(* IEC 61131-3 sources: Lasal-MCP/examples/SampleSource/LASALScreenAdvancedSolution/LASALScreenAdvancedSolution/LASALScreenAdvacnedSolution/Stations/MachineControl/MachineControl/Class/VaranManager (part 4) *)

      //look in all peripheral sync outs
      for i := 1 to VM_MAX_SYNC_OUTS - 1 do

        //look if sync out id is correct
        if ( p_SyncOut^.ucSyncOutID = VM_SYNC_OUT_ID ) then

          //if it is right pll for right manager number (first is vor VaranManager number 0, second for VaranManager number 1, ....)
          if ( ud_counter = 0 ) then
            exit;					//we found right sync out --> exit
          end_if;
          ud_counter -= 1;			//we find one for lower VaranManager number
        end_if;

        //get pointer to next sync out
        p_SyncOut += sizeof ( LSL_VARANPLLSYNCOUT );

        //if we searched all sync outs set VaranManager off
        if ( i = VM_MAX_SYNC_OUTS - 1 ) then
          p_SyncOut := NIL;
          State 		:= _NotInitialized;
          ManagerOn	:= 0;
          return;
        end_if;
      end_for;

      //disable varan manager sync out
      p_SyncOut^.ucControlStatus := 0;
    end_if;

  else // if b_PayloadSupport ****************************************************************************

    // if there is no VARAN Interface available, we would crash at the call
    if pVaran = NIL then
      sd_retval := VARANMANAGER_DRIVER_NOT_EXISTS;
      return;
    end_if;

      //-----------------------------------------------------------------------------------------------
    //get manager node info from os
    ManagerNodeString := 0;

    //call OS - function (must be OS-funciton because of error handling)
    sd_retval := VARAN_iGetNodeInfo	( uiManager	:= VaranManagerNr
                                    , pucNode	  := #ManagerNodeString
                                    , pNodeInfo	:= #p_NodeInfo
                                    );

    if	( sd_retval <> VARANMANAGER_OK
      | p_NodeInfo = NIL
      )
    then
      State := _NoHardware;
      return;
    end_if;

      // get release of FPGA
    Release := p_NodeInfo^.ucFPGAVersion;

    //-----------------------------------------------------------------------------------------------
    //get Manager structure
    sd_retval := VARAN_iGetManagerControl	( uiManager := VaranManagerNr
                                          , pvCB 		  := ( #p_ManagerStructure )$^PLSL_CONTROLBLOCK
                                          , pvPLL		  := ( #p_ManagerPll )$^PLSL_VARANPLL
                                          );

    //look for an error
    if	( sd_retval 			<> 	VARANMANAGER_OK
      | p_ManagerStructure	=	NIL
      | p_ManagerPll			= 	NIL
      )
    then
      State 		:= _NotInitialized;
      ManagerOn	:= 0;
      return;
    end_if;

    //look for right sync out pointer
    p_SyncOut := #p_ManagerPll^.sSynOutPeripheral1;
    ud_Counter := VaranManagerNr;

    //look in all peripheral sync outs
    for i := 1 to VM_MAX_SYNC_OUTS - 1 do

      //look if sync out id is correct
      if ( p_SyncOut^.ucSyncOutID = VM_SYNC_OUT_ID ) then

        //if it is right pll for right manager number (first is for VaranManager number 0, second for VaranManager number 1, ....)
        if ( ud_counter = 0 ) then
          exit;					//we found right sync out --> exit
        end_if;
        ud_counter -= 1;			//we find one for lower VaranManager number
      end_if;

      //get pointer to next sync out
      p_SyncOut += sizeof ( LSL_VARANPLLSYNCOUT );

      //if we searched all sync outs set VaranManager off
      if ( i = VM_MAX_SYNC_OUTS - 1 ) then
        p_SyncOut := NIL;
        State 		:= _NotInitialized;
        ManagerOn	:= 0;
        return;
      end_if;
    end_for;

    //disable varan manager sync out
    p_SyncOut^.ucControlStatus := 0;

    //set required bit on (for varan error in init (os set bit in function InitApp) later)
    p_ManagerStructure^.ucTCEnable := p_ManagerStructure^.ucTCEnable or 16#80;

    //Get ISO start Time
    GetISOStartTime();

    p_ManagerStructure^.uiIsoStartPoint := VaranManagerTime * IsoStartPoint / 100;

  end_if; // if b_PayloadSupport ****************************************************************************

  // get maintimer in ns to compare with varan times
  MainTimer := _ClockTicks * 1000;

  //look if VaranManagerTime is a multiple of maintimer (maintimer has to be always less or equal the varan time)
  if ( VaranManagerTime mod MainTimer <> 0 ) then
    //Log entry
#ifdef HWC_LogValue2
    HWC_LogValue2(this, "@064A (VaranManager::FirstInit) VaranManagerTime ({0}) is not a multiple of MainTimer ({1})!", VaranManagerTime, MainTimer);
#endif

    State 		:= _NotInitialized;
    ManagerOn	:= 0;
    return;
  end_if;

//------------------------------------------------------------ Client Instructions --------------------------------------------------------|
//                                                                                                                                         V
  if ( IsAlsoClient ) then

    if b_PayloadSupport &
       pMultiVaran^.udVersion >= VM_MULTIVARAN_VERSION_FULL_PAYLOAD_AVAILABLE  then
      sd_retval := MULTI_VARAN_iGetNodeProperty(  hNodeHandle       := vmNodeHandle
                                                , udPropertyId      := VC_OPT_PROP_BUFFER_ADDRESS_ISO // = Offset 0 in p_ManagerClientSpace
                                                , pudPropertyValue  := (#p_ManagerClientSpace)$^UDINT );

    elsif ( _RTOSVersion >= 16#11DA ) & pVaran then

      //Schnittstelle vom OS holen!!!!!!
      sd_retval := VARAN_iGetManagerClientAddress	( uiManager		:= VaranManagerNr
                                                  , uiType		  := 0
                                                  , puiAddress	:= ( #p_ManagerClientSpace )$^UDINT
                                                  );
    end_if;

    //check if function is available
    if ( sd_retval <> VARANMANAGER_OK | p_ManagerClientSpace = NIL ) then

      IsAlsoClient := 0;

#ifdef HWC_LogError
      HWC_LogError(this, "@0654 (VaranManager::FirstInit) Client - Function not available but activated! (at least OS - Version 1.1.217 required)");
#endif
    else
      TriggerClientWD             := TRUE;
      bEnableManagerWithNoModules := TRUE; // activate, to ensure varan-client functionality if no varan clients are connected to the manager.
      sd_retval                   := InitMulDivVMC();

      //look for an error
      if ( sd_retval <> 0 ) then
        ManagerOn	:= 0;
        return;
      end_if;
    end_if;

  end_if;

//------------------------------------------------------------ Client Instructions --------------------------------------------------------^
//                                                                                                                                         |

  //get system periode time
  if b_PayloadSupport &
     pMultiVaran^.udVersion >= VM_MULTIVARAN_VERSION_FULL_PAYLOAD_AVAILABLE  then

    if MULTI_VARAN_iGetNodeProperty( hNodeHandle       := vmNodeHandle
                                , udPropertyId      := VM_PROP_PLL_SYSTEM_PERIOD_TIME
                                , pudPropertyValue  := #ud_SystemPeriod
                                ) <> VARANMANAGER_OK then

#ifdef HWC_LogError
      HWC_LogError(this,"@01A1 (VaranManager::FirstInit) Failed to get PLL System period time");
#endif

      State 		:= _NotInitialized;
      ManagerOn	:= 0;
      return;
    else
    ud_SystemPeriod *= 10;
    end_if;

  else
    ud_SystemPeriod := ( ( p_ManagerPll^.aucPeriod )$UDINT and 16#FF_FFFF ) * 10;
  end_if;

  //look if VaranManager is a multiple of system periode
  if ( VaranManagerTime mod ud_SystemPeriod <> 0 ) &
     ( ud_SystemPeriod mod VaranManagerTime <> 0 ) then
    IF ( _firstscan = TRUE ) THEN
      //Log entry
#ifdef HWC_LogValue2
      HWC_LogValue2(this, "@065E (VaranManager::FirstInit) VaranManagerTime ({0}) is not a multiple of System Period Time ({1})!", VaranManagerTime, ud_SystemPeriod);
#endif

    END_IF;
    State 		:= _NotInitialized;
    ManagerOn	:= 0;
    return;
  end_if;

  if ( IsAlsoClient = 0 ) then

    //-----------------------------------------------------------------------------------------------
    //set sync out signal for peripherie sync out
    p_SyncOut^.ucPeriodMultiplier 	:= TO_USINT( VaranManagerTime / ud_SystemPeriod );
  end_if;

  //-----------------------------------------------------------------------------------------------
  //Write sync out, cannot directly be written with payload support
  if b_PayloadSupport &
     pMultiVaran^.udVersion >= VM_MULTIVARAN_VERSION_GET_SYSTEM_PROPERTY_AVAILABLE  then

    sd_retval := MULTI_VARAN_ICONFIGUREPLLSYNCOUT( hManagerNodeHandle    := vmNodeHandle
                                    , udSyncOutId           := VM_SYNC_OUT_ID
                                    , udPeriodMultiplier    := p_SyncOut^.ucPeriodMultiplier
                                    , udFrameCountThreshold := p_SyncOut^.ucFrameCountThreshold
                                    , udControlStatus       := p_SyncOut^.ucControlStatus
                                    );
  end_if;

  //-----------------------------------------------------------------------------------------------
  //set function list for controlling class
  s_VMFunctions.p_This		                := this;
  s_VMFunctions.ud_VaranTime	            := VaranManagerTime;
  s_VMFunctions.b_IsAlsoClient            := to_bool(IsAlsoClient);
  s_VMFunctions.ud_SuperiorTime           := SuperiorSystemTime;
  s_VMFunctions.SafetyManagerThisPointer  := #SafetyManagerThis;

  CoreSelect := CoreSelect.Read();

  //Check for correct setting
  if CoreSelect < TASK_SELECT_CORE0 | CoreSelect > TASK_SELECT_COREMAX then

#ifdef HWC_LogValue2
      HWC_LogValue2(this, "@01A2 (VaranManager::FirstInit) Client CoreSelect is invalid. Max Value: 0x{0}, Set value: 0x{1}",TASK_SELECT_COREMAX,CoreSelect$UDINT);
#endif

    state := _InvalidConfguration;
    ManagerOn := 0;
    return;
  end_if;

  //send info to HwControl class
#ifdef CMD_LOGIN_VARANMANAGER

    MyPara.uiCmd := CMD_LOGIN_VARANMANAGER;
    MyPara.aPara[0] := VaranManagerNr$DINT;               //Number of the VaranManager
    MyPara.aPara[1] := (#s_VMFunctions)$DINT;             //Pointer to function list
    MyPara.aPara[2] := CoreSelect$DINT;                   //Selection on which core the manager should be called (0 ... Core 0, 1 ... Core 1)
    MyPara.aPara[3] := ( VaranManagerTime / 1000 )$DINT;  //ud_RtTime_us

    //Always set cyclic to 1ms, except we have a maintimer which is greater than 1ms, then set it to maintimer (to have the same behaviour like the old system)
    if _ClockTicks > 1000 then
      udTempCyTime := _ClockTicks;
    else
      udTempCyTime := 1000;
    end_if;

    MyPara.aPara[4] := udTempCyTime$DINT;  //ud_CyTime_us

    To_HwControl.NewInst(pPara:=#MyPara, pResult:=#MyResult);

    sd_retval := MyResult.aData[0]$DINT;

#else

    if CoreSelect > TASK_SELECT_CORE0 then
#ifdef HWC_LogError
      HWC_LogError(this, "@01A3 (VaranManager::FirstInit) Need newer version of HwControl.h Headerfile. CoreSelect is not supported. Varanmanager will be called from the first CPU-core.");
#endif
      state := _InvalidConfguration;
      ManagerOn := 0;
      return;
    end_if;

    sd_retval := To_HwControl.AddVaranManager	( ud_manager_number	:= VaranManagerNr
                                              , p_function_list	  := #s_VMFunctions
                                              );
#endif

  //look for an error
  if ( sd_retval <> 0 ) then

#ifdef HWC_LogValue1
      HWC_LogValue1(this, "@01A4 (VaranManager::FirstInit) Failed to add VaranManager to HWControl. ErrorCode: 0x{0}!",sd_retval$UDINT);
#endif

    State 		:= _NotInitialized;
    ManagerOn	:= 0;
    return;
  end_if;

  //Check if we have the ability to give the OS the information which VaranManager runs on which processor core
  //The processing of the interrupts affecting this varanmanager also takes place on the same processor core as the realtime/cyclic of the hardware classes
  //*******************************************************************************************************
  if b_PayloadSupport & pMultiVaran^.udVersion >= VM_MULTIVARAN_VERSION_SET_CORESELECT_INFO_AVAILABLE then

    //Property ID of CoreSelect
    nodeProperty[0].udPropertyId    := VM_PROP_CORE_NUMBER;

    //Set Coreselect (0 ... first core, 1 ... second core, ...)
    nodeProperty[0].udPropertyValue := CoreSelect$UDINT;

    sd_retval := MULTI_VARAN_iSetNodeProperties( hNodeHandle           := vmNodeHandle
                                               , udPropertyCount       := 1
                                               , psPropertyValuePairs  := #nodeProperty[0]
                                               );

    if sd_retval <> VARANMANAGER_OK then
    #ifdef HWC_LogError
      HWC_LogError(this, "@04A9 (VaranManager::FirstInit) Failed to set core select information for OS! (VM_PROP_CORE_NUMBER)");
    #endif

      State 		:= _NotInitialized;
      ManagerOn	:= 0;
      return;
    end_if;
  end_if;
  //*******************************************************************************************************

  //-----------------------------------------------------------------------------------------------
  //install callback function for Timslice and watchdog error
  sd_retval := SetObjectCallback	( p_us_position_info	:= NIL
                                  , ud_action_ptr			  := ( #Varan_CallBack() )$UDINT
                                  , ud_thisp				    := this$UDINT
                                  , sd_required			    := 0
                                  );

  //look if an error occurs
  if ( sd_retval <> VARANMANAGER_OK ) then

#ifdef HWC_LogValue1
      HWC_LogValue1(this, "@065E (VaranManager::FirstInit) Failed to install callback function for Timeslice and watchdog error. Errorcode: 0x{0}",sd_retval$UDINT);
#endif

    State 		  := _CallBackError;
    ManagerOn 	:= 0;
    return;
  end_if;

  //-----------------------------------------------------------------------------------------------
  //Semaphore for direct accesses

  _strcpy(dest:=#aStrSemaphore[0], src:="VM_DA_SEMA_");

  ASCII_BIN1.Bin2Ascii(pt:=#astrVaranManagerNr[0], value:=to_dint(VaranManagerNr), format:=16#800);
  _strcat(dest:=#aStrSemaphore[0], src:=#aStrVaranManagerNr[0]);

  p_SemaHandle := To_Multitask.CreateSemaphore( MTSEMATYPE_RESOURCE, 1, 0, #aStrSemaphore[0] );
  if( p_SemaHandle = NIL )then
    State 		:= _NotInitialized;
    ManagerOn	:= 0;
#ifdef HWC_LogError
    HWC_LogError(this, "@0668 (VaranManager::FirstInit) Unable to create semaphore for async access!");
#endif
  end_if;

  //-----------------------------------------------------------------------------------------------
  if b_PayloadSupport &
     pMultiVaran^.udVersion >= VM_MULTIVARAN_VERSION_FULL_PAYLOAD_AVAILABLE  then
    // p_SyncAndWdDO p_SyncData are handled by OS when there is Payload Support

    //set periode of varan system
    nodeProperty[0].udPropertyId     := VM_PROP_PLL_SYSTEM_PERIOD_TIME;  // Also sets p_SyncData^.ui_Periode
    nodeProperty[0].udPropertyValue  := VaranManagerTime / 10 ;

    MULTI_VARAN_iSetNodeProperties( hNodeHandle           := vmNodeHandle
                                  , udPropertyCount       := 1
                                  , psPropertyValuePairs  := #nodeProperty[0]);

  else
    //get data of Sync and Watchdog DO
    sd_retval := VARAN_iGetSyncAndWdDO	( uiManager	:= VaranManagerNr
                                        , pvDO		  := #p_SyncAndWdDO
                                        , pvData	  := #p_SyncData$pvoid
                                        );

    //look for an error
    if	(( sd_retval <> VARANMANAGER_OK ) &
         ( s_VaranManagerSettings.us_InitCounter >= 10 )) then
      State 		:= _NotInitialized;
      ManagerOn	:= 0;
      return;
    end_if;

    //set periode of varan system
    p_SyncData^.ui_Periode := TO_UINT(  VaranManagerTime / 10 );				  //in 10ns steps
    p_SyncData^.us_Periode := TO_USINT( VaranManagerTime / 10 SHR 16 );		//in 10ns steps
  end_if;

  //set timemark for triggering watchdog
  s_VaranManagerSettings.ud_WatchdogTimemark := ops.tAbsolute - VM_WATCHDOG_TRIGGER_TIME;

END_FUNCTION

FUNCTION VaranManager::ExtendModuleList
  VAR_OUTPUT
    sd_retval   : DINT;
  END_VAR

  sd_retval := VARANMANAGER_OK;
    //--------------------------------------------------------------------------------------------------------------------
  //set right max handle
  s_ModuleList.ud_MaxModules += VM_EXTEND_HANDLES;

  //realloc memory for list
  s_ModuleList.p_ModuleList$^void := To_StdLib.ReAlloc	( mptr 		  := s_ModuleList.p_ModuleList
                                                        , newsize 	:= s_ModuleList.ud_MaxModules * sizeof( p_VaranBase )
                                                        );

  //look if we got memory for our Handle list
  if ( s_ModuleList.p_ModuleList ) then

    //set new memory to 0
    To_StdLib.MemSet( dest 	:= s_ModuleList.p_ModuleList + ( s_ModuleList.ud_MaxModules - VM_EXTEND_HANDLES ) * sizeof( p_VaranBase )
                    , value := 0
                    , size 	:= VM_EXTEND_HANDLES * sizeof( p_VaranBase )
                    );

  else
    //if not give out a TRACE
    sd_retval := VARANMANAGER_NO_MEM;

    //Log entry
#ifdef HWC_LogValue1
    HWC_LogValue1(this, "@0027 (VaranManager::ExtendModuleList) No Memory for Varan Manager available! (Extend Module List: {0})", s_ModuleList.ud_MaxModules);
#endif
  end_if;

  s_ModuleList.p_PositionList$^void := To_StdLib.ReAlloc( mptr     := s_ModuleList.p_PositionList
                                                        , newsize  := s_ModuleList.ud_MaxModules * sizeof (pVoid)
                                                        );

  //look if we got memory for our Handle list
  if ( s_ModuleList.p_PositionList ) then

    //set new memory to 0
    To_StdLib.MemSet( dest 	:= s_ModuleList.p_PositionList + ( s_ModuleList.ud_MaxModules - VM_EXTEND_HANDLES ) * sizeof( pVoid )
                    , value := 0
                    , size 	:= VM_EXTEND_HANDLES * sizeof(pVoid )
                    );

  else
    //if not give out a TRACE
    sd_retval := VARANMANAGER_NO_MEM;

    //Log entry
#ifdef HWC_LogValue1
    HWC_LogValue1(this, "@0028 (VaranManager::ExtendModuleList) No Memory for Varan Manager available! (Extend Position List: {0})", s_ModuleList.ud_MaxModules);
#endif
  end_if;

END_FUNCTION

FUNCTION GLOBAL VaranManager::CreateMutex
  VAR_INPUT
    MutexName 	      : ^CHAR;
    pThis 	          : ^VirtualBase;
  END_VAR
  VAR_OUTPUT
    pv_RetMutex 	    : pVoid;
  END_VAR
  VAR
    str_ObjName       : array[0..255] of char;
    str_ObjNamePart1  : array[0..VARAN_MUTEX_NAME_MAX_LENGTH-1] of char;
    str_ObjNamePart2  : array[0..VARAN_MUTEX_NAME_END_LENGTH] of char; // +1 for 0 Termination
    str_CombinedName  : array[0..VARAN_MUTEX_NAME_MAX_LENGTH-1] of char;
    str_this          : array[0..11] of char; // 2 byty %m, 8 byte Address, 1 byte for 0 Termination

    ud_LenObjName     : UDINT;
    ud_LenStr         : UDINT;
    ud_SepLenStr      : UDINT;
    ud_LenCombObjName : UDINT;
    ud_LenThis        : UDINT;

  END_VAR

  pv_RetMutex := Nil; // Error OS_CILGetv failed

  if pThis = nil then
    pthis := this;
  end_if;

  if (mt_api = nil) then
    if(OS_CILGet("LSL_MULTITASK", #mt_api$void)) THEN
      mt_api := NIL;
    end_if;
  end_if;

  if mt_api then

    _memset(dest:=#str_ObjName[0],      usByte:=0, cntr:=sizeof(str_ObjName)      );
    _memset(dest:=#str_ObjNamePart1[0], usByte:=0, cntr:=sizeof(str_ObjNamePart1) );
    _memset(dest:=#str_ObjNamePart2[0], usByte:=0, cntr:=sizeof(str_ObjNamePart2) );
    _memset(dest:=#str_CombinedName[0], usByte:=0, cntr:=sizeof(str_CombinedName) );
    _memset(dest:=#str_this[0],         usByte:=0, cntr:=sizeof(str_this)         );

    ud_LenStr := _strlen(MutexName);

    ud_SepLenStr := _strlen(VARAN_STR_MUTEX_NAME_SEPERATOR);
    ud_LenObjName := _GetObjName(pThis:=pthis, pName:=#str_ObjName[0]);

    if (ud_LenStr < VARAN_MUTEX_NAME_MAX_LENGTH) then
      _strcpy(dest:=#str_CombinedName[0], src:=MutexName);
    else
      _strncpy(dest:=#str_CombinedName[0], src:=MutexName, max:=VARAN_MUTEX_NAME_MAX_LENGTH-1);
    end_if;

    if (ud_LenObjName + ud_LenStr) < VARAN_MUTEX_NAME_MAX_LENGTH then
      _strcat(dest:=#str_CombinedName[0], src:=#str_ObjName[0]);
    else
      _strncpy(dest:=#str_ObjNamePart1[0], src:= #str_ObjName[0], max:= VARAN_MUTEX_NAME_MAX_LENGTH - ud_LenStr - ud_SepLenStr - VARAN_MUTEX_NAME_END_LENGTH - 1);    // Copy Beginning of str_ObjName
      _strncpy(dest:=#str_ObjNamePart2[0], src:= #str_ObjName[ud_LenObjName-VARAN_MUTEX_NAME_END_LENGTH-1], max:=VARAN_MUTEX_NAME_END_LENGTH);  // Copy Last MUTEX_NAME_END_LENGTH Char of str_ObjName

      // Put the Mutex String together
      _strcat(dest:=#str_CombinedName[0], src:= #str_ObjNamePart1[0]);
      _strcat(dest:=#str_CombinedName[0], src:= VARAN_STR_MUTEX_NAME_SEPERATOR);
      _strcat(dest:=#str_CombinedName[0], src:= #str_ObjNamePart2[0]);
    end_if;

    pv_RetMutex := OS_MT_CreateSemaphore(MTSEMATYPE_MUTEX, 1, 0, #str_CombinedName[0]);

    if pv_RetMutex = nil then

      // If Create Mutex failed: Insert the this pointer into the string
      ud_LenCombObjName := _strlen(#str_CombinedName[0]);

      str_this[0] := '%';
      str_this[1] := 'm';
      _itoa(udNumber:=pthis$UDINT, pString:=#str_this[2]);
      ud_LenThis  := _strlen(src:=#str_this[0]);

      _strcpy(dest:=#str_CombinedName[ud_LenCombObjName-ud_LenThis], src:=#str_this[0]);

      pv_RetMutex := OS_MT_CreateSemaphore(MTSEMATYPE_MUTEX, 1, 0, #str_CombinedName[0]);

    end_if;

  end_if;

END_FUNCTION

FUNCTION GLOBAL VaranManager::MutexStart
  VAR_INPUT
    pMutex 	: pVoid;
  END_VAR

  if(pMutex <> NIL) then
    OS_MT_WAIT(pMutex);
  end_if;

END_FUNCTION

FUNCTION GLOBAL VaranManager::MutexStop
  VAR_INPUT
    pMutex 	: pVoid;
  END_VAR

  if(pMutex <> NIL) then
    OS_MT_SIGNAL(pMutex);
  end_if;

END_FUNCTION

FUNCTION VIRTUAL GLOBAL VaranManager::Control::NewInst
  VAR_INPUT
    pPara 	                  : ^CmdStruct;
    pResult 	                : ^Results;
  END_VAR
  VAR_OUTPUT
    ret_code 	                : IprStates;
  END_VAR
  VAR
    p_paraAddDO               : ^t_VM_CMD_AddDO;
    p_paraMovDO               : ^t_VM_CMD_AddMovDo;
    p_paraGetPointers         : ^t_VM_CMD_GetDataPointers;
    p_paraGetModuleHandel     : ^t_VM_CMD_GetModuleHandle;
    PostInitRetcode           : iprStates;
    pHelpPostInit             : ^t_s_PostInitList;
    i                         : UINT;
    pHelp                     : ^void;  // This pointer to call newinst
    // local variables for the Requested HWTString
    pStr_HWTRequested         : ^CHAR;
    ui_HWTRequestedLength     : UINT;
    us_HWTRequestedCurrIndex  : USINT;
    i_Req                     : UINT;
    // local variables for HWTStrings in the VM
    pStr_HWTVM                : ^CHAR;
    us_HWTVMLength            : USINT;
    i_VM                      : USINT;
    ud_ModuleIndex            : UDINT;
    b_ModuleFound             : BOOL;
    // local variables to safe currently found module
    pStr_HWTVMCurrent         : ^CHAR;
    ud_ModuleIndexCurrent     : UDINT;
    TempArray                 : ARRAY [0..SERNO_STRING_SIZE-1] OF USINT;
    a_HelpArray               : ARRAY[0..99] OF CHAR;
	  ud_StrSize                : UDINT;
    ud_MaxStrSize             : UDINT;
    sSPIIDHeader              : t_s_SPIListHeader;

    MyPara                    : CmdStruct;
    MyResult                  : results;

    //local variables for dummy mux callback
    sd_retval                 : DINT;
  END_VAR

  ret_code := READY;  // Overwritten on error

  CASE pPara^.uiCmd OF
//**********************************************************************************************************************************************************
    CMD_POST_INIT_CALL: // call from hwcontrol
      // Check Loader Version if function is supported
      if ops.uiLoaderVersion$UINT >= VM_POST_INIT_AVAILABLE then
        bPostInitActive := TRUE;

#ifdef _LSL_TARGETARCH_ARM  // IO Image only needed for ARM  CPUs
#ifdef VARAN_iSetOutputImage
        // the image is not copied from the shadow ram to the VM DPRAM so far => copy it
        if (b_IOImageWritten = FALSE) & b_IOImage then
          VARAN_iSetOutputImage(VaranManagerNr, VARAN_DOL_ASY);
          b_IOImageWritten := TRUE;
        end_if;
#endif
#endif

        // we wait here until the initialisation of the Varan Rt and the SDIAS Clients has been finished
        CyWork(0);

        if bPostInitModulesReady then

          MyPara.uiCmd := CMD_GET_SUPPORTED_FEATURES;

          //Check if post init done cmd will be called from hwcontrol
          To_HwControl.NewInst(pPara:=#MyPara, pResult:=#MyResult);
          if MyResult.aData$t_HWC_SupportedFeatureBits1.PostInitDoneCmdCalled = FALSE then
            bPostInitActive := FALSE;
          end_if;

          ret_code := READY;
        else
          ret_code := BUSY;
        end_if;
      else
        // Should be impossible as we never request a Postinit if the Loader version is incorrect.
#ifdef HWC_LogError
        HWC_LogError(this, "@01A5 (VaranManager::Control::NewInst) CMD_POST_INIT_CALL not supported with current Loader. Loader Version >= 02.02.137 is required");
#endif
        ret_code := ERROR;
      end_if;

//**********************************************************************************************************************************************************
    CMD_POST_INIT_RT_SYNC:
      // check if all modules are ready
      if WaitForSyncSendObjectsCnt then
        CyWork(0);

        ret_code := BUSY;
      end_if;

//**********************************************************************************************************************************************************
    CMD_POST_INIT_RT_READY:
      // check post init modules
      if PostInitModuleCnt then
        pHelpPostInit := #aPostInitList[0];
        for i := 0 to PostInitModuleCnt - 1 do

          //call class, if it's still not ready
          if pHelpPostInit^.p_This then
            PostInitRetcode := pHelpPostInit^.p_This^.NewInst(pPara, pResult);

            // only overwrite the ready returncode if the returncode from the post init objects is different to it
            if PostInitRetcode <> READY then
              ret_code := PostInitRetcode;
            end_if;
          end_if;

          // set pointer on next this pointer
          pHelpPostInit += sizeof(t_s_PostInitList);
        end_for;
      end_if;

      // if manager is disabled => return error
      if ManagerOn = 0 then
        ret_code := ERROR;

      // if we're not ready, return busy
      elsif us_RtStep <> _RtWork then
        ret_code := BUSY;

      elsif ret_code = READY then
        // everything ready
        b_PostInitRtSyncReady := TRUE;
      end_if;

//**********************************************************************************************************************************************************
    CMD_SET_POSTINIT_DONE:  //call from hwcontrol

      //HwControl Postinit phase now finished.
      bPostInitActive := FALSE;

//**********************************************************************************************************************************************************
    CMD_FORCE_POST_INIT_END:  // call from hwcontrol
      // HWControl has run into timeout and has ended the Post Init Phase
      // This call informs the VM thats the Phase has ended.
      bPostInitActive := FALSE;

      //Check if this manager is the reason for the timeout, show it on server
      if ManagerOn <> 1 then
        State := _TimeoutInInit;
      end_if;

//**********************************************************************************************************************************************************
    CMD_POST_INIT_DO_SORT:    // call from hwcontrol
      // sort safety DOs if there is more than 1
      if pPriorityList & pPriorityList^.pNext &
        b_PayloadSupport = false then     // OS Handles Priorities of DO if b_PayloadSupport = true

        SortCmdsByPriority();

#ifdef _LSL_TARGETARCH_ARM  // IO Image only needed for ARM  CPUs
#ifdef VARAN_iSetOutputImage
        // Varandata has to be written once after sorting the DOs
        if b_IOImage then
          VARAN_iSetOutputImage(VaranManagerNr, VARAN_DOL_ISO);
        end_if;
      else
        // Varandata has to be written once after adding the DOs even without sorting anything because we need the shadow RAM image in the VM DPRAM)
        if b_IOImage then
          VARAN_iSetOutputImage(VaranManagerNr, VARAN_DOL_ISO);
        end_if;
#endif
#endif
      end_if;

//**********************************************************************************************************************************************************
    CMD_GET_HARDWARE_TREE_ENTRY:

      pHelp                     := nil;  // This pointer to call newinst
      // local variables for the Requested HWTString
      ui_HWTRequestedLength     := 0;
      us_HWTRequestedCurrIndex  := 0;
      i_Req                     := 0;
      // local variables for HWTStrings in the VM
      pStr_HWTVM                := NIL;
      us_HWTVMLength            := 0;
      i_VM                      := 0;
      ud_ModuleIndex            := 0;
      b_ModuleFound             := FALSE;

      // local variables to safe currently found module
      pStr_HWTVMCurrent         := NIL;
      ud_ModuleIndexCurrent     := 0;

      ret_code := ERROR;
      pResult^.aData[0]$t_HWCGetHardwareTreeEntryOut.retcode := _HWC_RETVAL_ERROR_VARAN_MODULE_NOT_FOUND;

      pStr_HWTRequested     := pPara^.aPara[0]$t_HWCGetHardwareDiagnosisIn.pStr_HardewareTreeEntry;

      //First HWT Path
      if pStr_HWTRequested = nil then

        ud_VaranPosition := VM_OBJECT_PATH;

        // Return String of the Varanmanger
        ret_code := READY;
        pResult^.aData$t_HWCGetHardwareTreeEntryOut.retcode := _HWC_RETVAL_OK_HWTSTR_RETURNED;
        pResult^.aData[0]$t_HWCGetHardwareTreeEntryOut.pStr_NextHardewareTreeEntry := (#ud_VaranPosition)$^CHAR;

      // Only possible for VM own HWT Path
      elsif (pStr_HWTRequested^$USINT = 2) then

        if pStr_HWTRequested^$UDINT = VM_OBJECT_PATH then

          if s_ModuleList.p_ModuleList^ then
            // Return first Module in list
            ret_code := s_ModuleList.p_ModuleList^$p_VaranBase^.NewInst(pPara,pResult);
          else
            // VM was found but there are no modules connected
            ret_code := READY;
            pResult^.aData[0]$t_HWCGetHardwareTreeEntryOut.retcode := _HWC_RETVAL_OK_MODULE_FOUND;
          end_if;
        end_if;

      else

        //Search for module
        ui_HWTRequestedLength     := (pStr_HWTRequested)$^UINT^ + 1;  //+1 because we compare the strings, 2 byte length
        us_HWTRequestedCurrIndex  := pPara^.aPara[0]$t_HWCGetHardwareDiagnosisIn.us_current_index;

        ud_ModuleIndex := 0;
        b_ModuleFound := FALSE;

        //loop over all modules
        while (ud_ModuleIndex < s_ModuleList.ud_NrOfModules) &
              (b_ModuleFound = FALSE) do

          pStr_HWTVM := (s_ModuleList.p_PositionList+ (ud_ModuleIndex * 4))^$^CHAR;  // 4 = SizeOf(^CHAR)

          if pStr_HWTVM  then
            us_HWTVMLength := pStr_HWTVM^;  //First byte is length

            i_Req := us_HWTRequestedCurrIndex;
            i_Vm  := 1;

            //Loop over strings
            while i_Req <= ui_HWTRequestedLength &
                  i_Vm  <= us_HWTVMLength do

              if (pStr_HWTRequested + i_Req)^ <> (pStr_HWTVM + i_Vm)^ then // Compare byte
                // Strings are not equal
                exit;
              end_if;

              i_Req += 1;
              i_VM  += 1;
            end_while;

            if (i_Req <= ui_HWTRequestedLength ) &                        // End of requested string was not reached
               (i_Vm = us_HWTVMLength + 1) &                              // And end of compared string reached
               ( (pStr_HWTRequested + i_Req)^ and HWT_ESCAPE_SEQU ) then  // Escape sequece found in Requested string

              b_ModuleFound := TRUE;

//              pPara^.aPara[0]$t_HWCGetHardwareDiagnosisIn.us_current_index   := i_Req$USINT;
//              pPara^.aPara[0]$t_HWCGetHardwareDiagnosisIn.us_current_length  := (ui_HWTRequestedLength - i_Req)$USINT;
              exit;
            end_if;

            if (i_Vm = us_HWTVMLength + 1) & (i_Req = ui_HWTRequestedLength + 1) then   // All Bytes and Length are equal
              b_ModuleFound := TRUE;

//              pPara^.aPara[0]$t_HWCGetHardwareDiagnosisIn.us_current_index  := i_Req$USINT - 1;  // -1 because we increased over max length at the end of the while loop
//              pPara^.aPara[0]$t_HWCGetHardwareDiagnosisIn.us_current_length := 1; // Last entry of string was reached, index points to last entry
              exit;
            end_if;

          end_if;

          ud_ModuleIndex += 1;  // Select next Module

        end_while;

        if b_ModuleFound then

          // Call module again incase it is an extension module
          pHelp     := s_ModuleList.p_ModuleList + sizeof(p_VaranBase) * ud_ModuleIndex;
          ret_code  := pHelp^$p_VaranBase^.NewInst(pPara,pResult);

          // Return if new HWT String was found
          if ret_code = READY &
             pResult^.aData[0]$t_HWCGetHardwareDiagnosisOut.retcode = _HWC_RETVAL_OK_HWTSTR_RETURNED then
            return;
          end_if;

          ud_ModuleIndex        += 1;  // Select next Module
          ud_ModuleIndexCurrent := ud_ModuleIndex;

          b_ModuleFound := TRUE;  // Only set to enter loop

          while (ud_ModuleIndexCurrent < s_ModuleList.ud_NrOfModules) &
                (b_ModuleFound = TRUE) do

            pStr_HWTVMCurrent := (s_ModuleList.p_PositionList+ (ud_ModuleIndexCurrent * 4))^$^CHAR ;  // 4 = SizeOf(^CHAR)

            if pStr_HWTVMCurrent then

              // Check if module has already been called (multiple entries in list)
              ud_ModuleIndex  := 0;
              b_ModuleFound   := FALSE;

              //loop over all modules to search for duplicates
              while (ud_ModuleIndex < ud_ModuleIndexCurrent &
                     b_ModuleFound = FALSE) do

                pStr_HWTVM := (s_ModuleList.p_PositionList+ (ud_ModuleIndex * 4))^$^CHAR ;  // 4 = SizeOf(^CHAR)

                if pStr_HWTVM then

                  // Compare string length
                  if pStr_HWTVMCurrent^ = pStr_HWTVM^ then

                    // Compare string content
                    if _memcmp( ptr1 := pStr_HWTVMCurrent + 1,
                                ptr2 := pStr_HWTVM +1,
                                cntr := pStr_HWTVMCurrent^) = 0 then

                      // Multiple entry, Check next Module
                      b_ModuleFound         := TRUE;
                      ud_ModuleIndexCurrent += 1;
                      exit;

                    end_if;
                  end_if;
                end_if;

                ud_ModuleIndex += 1;

              end_while;

              if b_ModuleFound = FALSE then
                exit; // Non duplicate entry
              end_if;

            else  // if pStr_HWTVMCurrent then
              ud_ModuleIndexCurrent += 1;
            end_if;

          end_while;

          if b_ModuleFound = FALSE then
            // Call Class
            pHelp     := s_ModuleList.p_ModuleList + sizeof(p_VaranBase) * ud_ModuleIndexCurrent;
            ret_code  := pHelp^$p_VaranBase^.NewInst(pPara,pResult);
          end_if;

        else
          pResult^.aData[0]$t_HWCGetHardwareDiagnosisOut.retcode := _HWC_RETVAL_ERROR_VARAN_MODULE_NOT_FOUND;
          ret_code := ERROR;
        end_if;

      end_if;

//**********************************************************************************************************************************************************
    CMD_GET_HARDWARE_DIAGNOSIS:

      pHelp                     := nil;  // This pointer to call newinst
      // local variables for the Requested HWTString
      ui_HWTRequestedLength     := 0;
      us_HWTRequestedCurrIndex  := 0;
      i_Req                     := 0;
      // local variables for HWTStrings in the VM
      pStr_HWTVM                := NIL;
      us_HWTVMLength            := 0;
      i_VM                      := 0;
      ud_ModuleIndex            := 0;
      b_ModuleFound             := FALSE;

      ret_code := ERROR;
      pResult^.aData[0]$t_HWCGetHardwareDiagnosisOut.retcode := _HWC_RETVAL_ERROR;

      pStr_HWTRequested     := pPara^.aPara[0]$t_HWCGetHardwareDiagnosisIn.pStr_HardewareTreeEntry;

      if pStr_HWTRequested then

        // Check for VM String
        if (pStr_HWTRequested)$^UINT^ = 2 then

          if (pStr_HWTRequested)$^UDINT^ = VM_OBJECT_PATH then

            TempArray[0] := 0;

            if this <> p_this then
              //Reset statemachine
              eSPISSW := _GetVendorName;
              //Save This pointer
              p_this := this;

              // Reset Flags
              bDiagnosisDataAvailableFlags.HWVersion   := FALSE;
              bDiagnosisDataAvailableFlags.VendorName  := FALSE;
              bDiagnosisDataAvailableFlags.DeviceName  := FALSE;
              bDiagnosisDataAvailableFlags.OrderingNo  := FALSE;
              bDiagnosisDataAvailableFlags.LicenseNo   := FALSE;
              bDiagnosisDataAvailableFlags.SerialNo    := FALSE;
            end_if;

            case eSPISSW of
            	_GetVendorName:
                ret_code$DINT := GetSPIDataFromID(  p_us_position_info  := #TempArray[0]
                                                  , udListID            := VM_SPI_VENDOR_NAME_ID
                                                  , pData               := #a_VendorName[0]
                                                  , udRequDataLength    := sizeof(a_VendorName)
                                                  , pIDHeader           := #sSPIIDHeader
                                                  );

                if ret_code = READY then

                  // Null Termination ----------------------------------------
                  ud_StrSize    := sSPIIDHeader.ListLength;
                  ud_MaxStrSize := sizeof(a_VendorName);

                  pResult^.aData[0]$t_HWCGetHardwareDiagnosisOut.pStr_VendorName                    := (#a_VendorName)$^CHAR; // Will be overwritten if this pointer is not equal

                  (pResult^.aData[0]$t_HWCGetHardwareDiagnosisOut.pStr_VendorName + ud_MaxStrSize)^ := 0;
                  if ud_StrSize < ud_MaxStrSize then
                    (pResult^.aData[0]$t_HWCGetHardwareDiagnosisOut.pStr_VendorName + ud_StrSize)^  := 0;
                  end_if;

                  bDiagnosisDataAvailableFlags.VendorName := TRUE;

                  eSPISSW := _GetSerialNo;
                  ret_code := BUSY;
                else
                  pResult^.aData[0]$t_HWCGetHardwareDiagnosisOut.retcode := _HWC_RETVAL_ERROR_VARAN_SPI_ACCESS_FAILED;
                  //set SSW to SPI Data Ready, because we return the values which are already in the HWK
                  eSPISSW := _SPIDataReady;
                  ret_code := BUSY;
                end_if;

              _GetSerialNo:
                ret_code$DINT := GetSPIDataFromID(  p_us_position_info  := #TempArray[0]
                                                  , udListID            := VM_SPI_SERIALNO_ID
                                                  , pData               := #a_SerialNo[0]
                                                  , udRequDataLength    := sizeof(a_SerialNo)
                                                  , pIDHeader           := #sSPIIDHeader
                                                  );

                if ret_code = READY then

                  // Null Termination ----------------------------------------
                  ud_StrSize    := sSPIIDHeader.ListLength;
                  ud_MaxStrSize := sizeof(a_SerialNo);

                  pResult^.aData[0]$t_HWCGetHardwareDiagnosisOut.pStr_SerialNo                    := (#a_SerialNo)$^CHAR; // Will be overwritten if this pointer is not equal

                  (pResult^.aData[0]$t_HWCGetHardwareDiagnosisOut.pStr_SerialNo + ud_MaxStrSize)^ := 0;
                  if ud_StrSize < ud_MaxStrSize then
                    (pResult^.aData[0]$t_HWCGetHardwareDiagnosisOut.pStr_SerialNo + ud_StrSize)^  := 0;
                  end_if;

                  bDiagnosisDataAvailableFlags.SerialNo := TRUE;

                  eSPISSW   := _GetDeviceName;
                  ret_code  := BUSY;
                else
                  pResult^.aData[0]$t_HWCGetHardwareDiagnosisOut.retcode := _HWC_RETVAL_ERROR_VARAN_SPI_ACCESS_FAILED;
                  //set SSW to SPI Data Ready, because we return the values which are already in the HWK
                  eSPISSW   := _SPIDataReady;
                  ret_code  := BUSY;
                end_if;

            	_GetDeviceName:
                ret_code$DINT := GetSPIDataFromID(  p_us_position_info  := #TempArray[0]
                                                  , udListID            := VM_SPI_DEVICE_NAME_ID
                                                  , pData               := #a_DeviceName[0]
                                                  , udRequDataLength    := sizeof(a_DeviceName)
                                                  , pIDHeader           := #sSPIIDHeader
                                                  );

                if ret_code = READY then

                  // Null Termination ----------------------------------------
                  ud_StrSize    := sSPIIDHeader.ListLength;
                  ud_MaxStrSize := sizeof(a_DeviceName);

                  pResult^.aData[0]$t_HWCGetHardwareDiagnosisOut.pStr_DeviceName                    := (#a_DeviceName)$^CHAR; // Will be overwritten if this pointer is not equal

                  (pResult^.aData[0]$t_HWCGetHardwareDiagnosisOut.pStr_DeviceName + ud_MaxStrSize)^ := 0;
                  if ud_StrSize < ud_MaxStrSize then
                    (pResult^.aData[0]$t_HWCGetHardwareDiagnosisOut.pStr_DeviceName + ud_StrSize)^  := 0;
                  end_if;

                  bDiagnosisDataAvailableFlags.DeviceName := TRUE;

                  eSPISSW   := _GetOrderingNo;
                  ret_code  := BUSY;
                else
                  pResult^.aData[0]$t_HWCGetHardwareDiagnosisOut.retcode := _HWC_RETVAL_ERROR_VARAN_SPI_ACCESS_FAILED;
                  //set SSW to SPI Data Ready, because we return the values which are already in the HWK
                  eSPISSW   := _SPIDataReady;
                  ret_code  := BUSY;
                end_if;

            	_GetOrderingNo:
                ret_code$DINT := GetSPIDataFromID(  p_us_position_info  := #TempArray[0]
                                                  , udListID            := VM_SPI_ORDERING_NO_ID
                                                  , pData               := #a_OrderingNo[0]
                                                  , udRequDataLength    := sizeof(a_OrderingNo)
                                                  , pIDHeader           := #sSPIIDHeader
                                                  );

                if ret_code = READY then

                  // Null Termination ----------------------------------------
                  ud_StrSize    := sSPIIDHeader.ListLength;
                  ud_MaxStrSize := sizeof(a_OrderingNo);

                  pResult^.aData[0]$t_HWCGetHardwareDiagnosisOut.pStr_OrderingNo                    := (#a_OrderingNo)$^CHAR; // Will be overwritten if this pointer is not equal

                  (pResult^.aData[0]$t_HWCGetHardwareDiagnosisOut.pStr_OrderingNo + ud_MaxStrSize)^ := 0;
                  if ud_StrSize < ud_MaxStrSize then
                    (pResult^.aData[0]$t_HWCGetHardwareDiagnosisOut.pStr_OrderingNo + ud_StrSize)^  := 0;
                  end_if;

                  bDiagnosisDataAvailableFlags.OrderingNo := TRUE;

                  eSPISSW   := _GetLicenseNoHWVersion;
                  ret_code  := BUSY;
                else
                  pResult^.aData[0]$t_HWCGetHardwareDiagnosisOut.retcode := _HWC_RETVAL_ERROR_VARAN_SPI_ACCESS_FAILED;
                  //set SSW to SPI Data Ready, because we return the values which are already in the HWK
                  eSPISSW   := _SPIDataReady;
                  ret_code  := BUSY;
                end_if;

            	_GetLicenseNoHWVersion:

                ret_code$DINT := GetSPIDataFromID(  p_us_position_info  := #TempArray[0]
                                                  , udListID            := VM_SPI_IDENTIFICATION_LIST
                                                  , pData               := #a_HelpArray[0]
                                                  , udRequDataLength    := sizeof(udHWVersion) + sizeof(udLicenseNo)
                                                  , pIDHeader           := #sSPIIDHeader
                                                  , udOffset            := 8
                                                  );

                udLicenseNo := a_HelpArray[0]$UDINT;
                udHWVersion := a_HelpArray[4]$UDINT;

                if ret_code = READY then
                  bDiagnosisDataAvailableFlags.LicenseNo := TRUE;
                  bDiagnosisDataAvailableFlags.HWVersion := TRUE;
                  eSPISSW   := _SPIDataReady;
                  ret_code  := BUSY;
                else
                  pResult^.aData[0]$t_HWCGetHardwareDiagnosisOut.retcode := _HWC_RETVAL_ERROR_VARAN_SPI_ACCESS_FAILED;
                  //set SSW to SPI Data Ready, because we return the values which are already in the HWK
                  eSPISSW   := _SPIDataReady;
                  ret_code  := BUSY;
                end_if;

            	_SPIDataReady:
                //Don't reset statemachine because if we have the same this pointer we don't have to make spi Accesses again
                //eSPISSW := _GetVendorName;

                //Data which is already in HWK available
                if p_NodeInfo then

                  pResult^.aData$t_HWCGetHardwareDiagnosisOut.hd_FPGAVersion      := to_udint(p_NodeInfo^.ucFPGAVersion);
                  pResult^.aData$t_HWCGetHardwareDiagnosisOut.ud_DeviceID         := to_udint(p_NodeInfo^.uiDeviceID);
                  pResult^.aData$t_HWCGetHardwareDiagnosisOut.ud_VendorID         := to_udint(p_NodeInfo^.uiVendorID);
                end_if;

                if bDiagnosisDataAvailableFlags.VendorName then
                  pResult^.aData[0]$t_HWCGetHardwareDiagnosisOut.pStr_VendorName  := (#a_VendorName)$^CHAR;
                end_if;

                if bDiagnosisDataAvailableFlags.HWVersion & bDiagnosisDataAvailableFlags.LicenseNo then
                  pResult^.aData[0]$t_HWCGetHardwareDiagnosisOut.hd_HWVersion     := udHWVersion;
                  pResult^.aData[0]$t_HWCGetHardwareDiagnosisOut.ud_LicenseNo     := udLicenseNo;
                end_if;

                if bDiagnosisDataAvailableFlags.DeviceName then
                  pResult^.aData[0]$t_HWCGetHardwareDiagnosisOut.pStr_DeviceName  := (#a_DeviceName)$^CHAR;
                end_if;

                if bDiagnosisDataAvailableFlags.OrderingNo then
                  pResult^.aData[0]$t_HWCGetHardwareDiagnosisOut.pStr_OrderingNo  := (#a_OrderingNo)$^CHAR;
                end_if;

                if bDiagnosisDataAvailableFlags.SerialNo then
                  pResult^.aData[0]$t_HWCGetHardwareDiagnosisOut.pStr_SerialNo    := (#a_SerialNo)$^CHAR;
                end_if;

                ret_code                                                          := READY;
                pResult^.aData[0]$t_HWCGetHardwareDiagnosisOut.retcode            := _HWC_RETVAL_OK;

            end_case;
          end_if;

          return;
        end_if;

        ui_HWTRequestedLength     := (pStr_HWTRequested)$^UINT^ + 1;  //+1 because we compare the strings, 2 byte length
        us_HWTRequestedCurrIndex  := pPara^.aPara[0]$t_HWCGetHardwareDiagnosisIn.us_current_index;

        ud_ModuleIndex := 0;
        b_ModuleFound := FALSE;

        //loop over all modules
        while (ud_ModuleIndex < s_ModuleList.ud_NrOfModules) &
              (b_ModuleFound = FALSE) do

          pStr_HWTVM := (s_ModuleList.p_PositionList+ (ud_ModuleIndex * 4))^$^CHAR ;  // 4 = SizeOf(^CHAR)

          if pStr_HWTVM  then
            us_HWTVMLength := pStr_HWTVM^;  //First byte is length

            i_Req := us_HWTRequestedCurrIndex;
            i_Vm  := 1;

            //Loop over strings
            while i_Req <= ui_HWTRequestedLength &
                  i_Vm  <= us_HWTVMLength do

              if (pStr_HWTRequested + i_Req)^ <> (pStr_HWTVM + i_Vm)^ then // Compare byte
                // Strings are not equal
                exit;
              end_if;

              i_Req += 1;
              i_VM  += 1;
            end_while;

            if (i_Req <= ui_HWTRequestedLength ) &                        // End of requested string was not reached
            (i_Vm = us_HWTVMLength + 1) &                                 // And end of compared string reached
               ( (pStr_HWTRequested + i_Req)^ and HWT_ESCAPE_SEQU ) then  // Escape sequece found in Requested string

              b_ModuleFound := TRUE;
              pPara^.aPara[0]$t_HWCGetHardwareDiagnosisIn.us_current_index   := i_Req$USINT;
              pPara^.aPara[0]$t_HWCGetHardwareDiagnosisIn.us_current_length  := (ui_HWTRequestedLength - i_Req)$USINT;
              exit;
            end_if;

            if (i_Vm = us_HWTVMLength + 1) & (i_Req = ui_HWTRequestedLength + 1) then   // All Bytes and Length are equal
              b_ModuleFound := TRUE;
              pPara^.aPara[0]$t_HWCGetHardwareDiagnosisIn.us_current_index  := i_Req$USINT - 1;  // -1 because we increased over max length at the end of the while loop
              pPara^.aPara[0]$t_HWCGetHardwareDiagnosisIn.us_current_length := 1; // Last entry of string was reached, index points to last entry
              exit;
            end_if;

          end_if;

          ud_ModuleIndex += 1;  // Select next Module

        end_while;

        if b_ModuleFound then
          // Call Class
          pHelp     := s_ModuleList.p_ModuleList + sizeof(p_VaranBase) * ud_ModuleIndex;
          ret_code  := pHelp^$p_VaranBase^.NewInst(pPara,pResult);
        else
          pResult^.aData[0]$t_HWCGetHardwareDiagnosisOut.retcode := _HWC_RETVAL_ERROR_VARAN_MODULE_NOT_FOUND;
          ret_code  := ERROR;
        end_if;

      end_if;

//**********************************************************************************************************************************************************
    VM_CMD_NEED_POST_INIT_CALL: // call from varan client
      // Check Loader Version if function is supported
      if ops.uiLoaderVersion$UINT >= VM_POST_INIT_AVAILABLE then

        // store this pointer of the module
        aPostInitList[PostInitModuleCnt].p_This := pPara^.aPara[0]$p_VaranBase;

        // remember if we have to wait for DOs to be created
        aPostInitList[PostInitModuleCnt].Settings := pPara^.aPara[1]$BSINT;
        if aPostInitList[PostInitModuleCnt].Settings.Wait4DOCreation then
          WaitForPostInitObjectsCnt += 1;
          if aPostInitList[PostInitModuleCnt].Settings.Wait4MoveDOCreation then
            WaitForPostInitMoveObjectsCnt += 1;
          end_if;
        end_if;

        // remember if we have to wait for the sync of this module
        if aPostInitList[PostInitModuleCnt].Settings.Wait4SyncSend then
          WaitForSyncSendObjectsCnt += 1;
        end_if;

        aPostInitList[PostInitModuleCnt].b_CallMe := TRUE;

        // return index for this module
        pResult^.uiLng          := 2;
        pResult^.aData[0]$UINT  := PostInitModuleCnt;

        // increase number of post init modules
        PostInitModuleCnt       += 1;

        // we're no longer ready with post init. we have to wait until all modules from the list are finished
        bPostInitModulesReady   := FALSE;
      else
#ifdef HWC_LogError
        HWC_LogError(this, "@01A6 (VaranManager::Control::NewInst) VM_CMD_NEED_POST_INIT_CALL not supported with current Loader. Loader Version >= 02.02.137 is required");
#endif
        ret_code := ERROR;
      end_if;

//**********************************************************************************************************************************************************
    VM_CMD_POST_INIT_FINISHED: // call from varan client
      // Check Loader Version if function is supported
      if ops.uiLoaderVersion$UINT >= VM_POST_INIT_AVAILABLE then

        // only relevant during last Init
        if PostInitModuleCnt then
          // check if it's a valid index
          if pPara^.aPara[1]$UINT < VM_MAX_POST_INIT_MODULES then
            // check if our local this pointer matches this object
            if pPara^.aPara[0]$p_VaranBase = aPostInitList[pPara^.aPara[1]$UINT].p_This then
              // increase number of ready objects
              PostInitModuleReadyCnt += 1;
//              aPostInitList[pPara^.aPara[1]$UINT].b_CallMe := FALSE;

              // check if it's an object we were waiting for
              if aPostInitList[pPara^.aPara[1]$UINT].Settings.Wait4DOCreation then
                aPostInitList[pPara^.aPara[1]$UINT].Settings.Wait4DOCreation := FALSE;

                if WaitForPostInitObjectsCnt then
                  WaitForPostInitObjectsCnt -= 1;
                else
#ifdef HWC_LogError
                  HWC_LogError(this, "@01A7 (VaranManager::Control::NewInst) There is already no more post init object to wait for! (VM_CMD_POST_INIT_FINISHED)");
#endif
                  ret_code := ERROR;
                end_if;
              end_if;

              // check if it's an object we were waiting for
              if aPostInitList[pPara^.aPara[1]$UINT].Settings.Wait4MoveDOCreation then
                aPostInitList[pPara^.aPara[1]$UINT].Settings.Wait4MoveDOCreation := FALSE;

                if WaitForPostInitMoveObjectsCnt then
                  WaitForPostInitMoveObjectsCnt -= 1;
                else
#ifdef HWC_LogError
                  HWC_LogError(this, "@01A8 (VaranManager::Control::NewInst) There is already no more post init object to wait for (create move DOs)! (VM_CMD_POST_INIT_FINISHED)");
#endif
                  ret_code := ERROR;
                end_if;
              end_if;

              // on last init we check if all modules which need to have finished their init
              if PostInitModuleReadyCnt = PostInitModuleCnt then
                bPostInitModulesReady := TRUE;
              end_if;
            else
#ifdef HWC_LogError
              HWC_LogError(this, "@01A9 (VaranManager::Control::NewInst) This pointer of post init module given doesn't match locally stored this pointer for this index!");
#endif
              ret_code := ERROR;
            end_if;
          else
#ifdef HWC_LogError
            HWC_LogError(this, "@01AA (VaranManager::Control::NewInst) Invalid index of post init module given!");
#endif
            ret_code := ERROR;
          end_if;
        else
#ifdef HWC_LogError
          HWC_LogError(this, "@01AB (VaranManager::Control::NewInst) More modules ready with last init than expected");
#endif
          ret_code := ERROR;
        end_if;
      else
#ifdef HWC_LogError
        HWC_LogError(this, "@01AC (VaranManager::Control::NewInst) VM_CMD_POST_INIT_FINISHED not supported with current Loader. Loader Version >= 02.02.137 is required");
#endif
        ret_code := ERROR;
      end_if;

//**********************************************************************************************************************************************************
    VM_CMD_IS_PAYLOAD_SUPPORTED:  // to get the status of PayloadSupport
      pResult^.aData[0]$BOOL := b_PayloadSupport;

//**********************************************************************************************************************************************************
    VM_CMD_DO_CREATION_FINISHED: // a post-init module is finished with creating DOs
      // Check Loader Version if function is supported
      if ops.uiLoaderVersion$UINT >= VM_POST_INIT_AVAILABLE then

        // only relevant during last Init
        if PostInitModuleCnt then
          // check if it's a valid index
          if pPara^.aPara[1]$UINT < VM_MAX_POST_INIT_MODULES then
            // check if our local this pointer matches this object
            if pPara^.aPara[0]$p_VaranBase = aPostInitList[pPara^.aPara[1]$UINT].p_This then
              // check if it's an object we were waiting for
              if aPostInitList[pPara^.aPara[1]$UINT].Settings.Wait4DOCreation then
                aPostInitList[pPara^.aPara[1]$UINT].Settings.Wait4DOCreation := FALSE;

                if WaitForPostInitObjectsCnt then
                  WaitForPostInitObjectsCnt -= 1;
                else
#ifdef HWC_LogError
                  HWC_LogError(this, "@01AD (VaranManager::Control::NewInst) There is already no more post init object to wait for!");
#endif
                  ret_code := ERROR;
                end_if;
              else
#ifdef HWC_LogError
                HWC_LogError(this, "@01AE (VaranManager::Control::NewInst) Module finished with DO creation, where  There is already no more post init object to wait for!");
#endif
                ret_code := ERROR;
              end_if;
            else
#ifdef HWC_LogError
              HWC_LogError(this, "@01A9 (VaranManager::Control::NewInst) This pointer of post init module given doesn't match locally stored this pointer for this index!");
#endif
              ret_code := ERROR;
            end_if;
          else
#ifdef HWC_LogError
            HWC_LogError(this, "@01AA (VaranManager::Control::NewInst) Invalid index of post init module given!");
#endif
            ret_code := ERROR;
          end_if;
        else
#ifdef HWC_LogError
          HWC_LogError(this, "@01AB (VaranManager::Control::NewInst) More modules ready with last init than expected");
#endif
          ret_code := ERROR;
        end_if;
      else
#ifdef HWC_LogError
        HWC_LogError(this, "@01AF (VaranManager::Control::NewInst) VM_CMD_DO_CREATION_FINISHED not supported with current Loader. Loader Version >= 02.02.137 is required");
#endif
        ret_code := ERROR;
      end_if;

//**********************************************************************************************************************************************************
    VM_CMD_MOVE_DO_CREATION_FINISHED:
      // Check Loader Version if function is supported
      if ops.uiLoaderVersion$UINT >= VM_POST_INIT_AVAILABLE then

        // only relevant during last Init
        if PostInitModuleCnt then
          // check if it's a valid index
          if pPara^.aPara[1]$UINT < VM_MAX_POST_INIT_MODULES then
            // check if our local this pointer matches this object
            if pPara^.aPara[0]$p_VaranBase = aPostInitList[pPara^.aPara[1]$UINT].p_This then
              // check if it's an object we were waiting for
              if aPostInitList[pPara^.aPara[1]$UINT].Settings.Wait4MoveDOCreation then
                aPostInitList[pPara^.aPara[1]$UINT].Settings.Wait4MoveDOCreation := FALSE;

                if WaitForPostInitMoveObjectsCnt then
                  WaitForPostInitMoveObjectsCnt -= 1;
                else
#ifdef HWC_LogError
                  HWC_LogError(this, "@01B0 (VaranManager::Control::NewInst) There is already no more post init object to wait for (create move DOs)!");
#endif
                  ret_code := ERROR;
                end_if;
              else
#ifdef HWC_LogError
                HWC_LogError(this, "@01B1 (VaranManager::Control::NewInst) Module finished with move DO creation, where  There is already no more post init object to wait for!");
#endif
                ret_code := ERROR;
              end_if;
            else
#ifdef HWC_LogError
              HWC_LogError(this, "@01B2 (VaranManager::Control::NewInst) This pointer of post init module given doesn't match locally stored this pointer for this index! (Move DOs)");
#endif
              ret_code := ERROR;
            end_if;
          else
#ifdef HWC_LogError
            HWC_LogError(this, "@01B3 (VaranManager::Control::NewInst) Invalid index of post init module given! (Move DOs)");
#endif
            ret_code := ERROR;
          end_if;
        else
#ifdef HWC_LogError
          HWC_LogError(this, "@01B4 (VaranManager::Control::NewInst) More modules ready with last init than expected (Move DOs)");
#endif
          ret_code := ERROR;
        end_if;
      else
#ifdef HWC_LogError
        HWC_LogError(this, "@01B5 (VaranManager::Control::NewInst) VM_CMD_MOVE_DO_CREATION_FINISHED not supported with current Loader. Loader Version >= 02.02.137 is required (Move DOs)");
#endif
        ret_code := ERROR;
      end_if;

//**********************************************************************************************************************************************************
    VM_CMD_DO_MEM_READY: // check if all post init objects are finished with creating DOs
      // if we're not in post init or the varan manager has finished waiting for post init objects => the DO memory is ready
      if WaitForPostInitObjectsCnt = 0 then
        pResult^.aData[4] := TRUE;
      else
        pResult^.aData[4] := FALSE;
      end_if;

//**********************************************************************************************************************************************************
    VM_CMD_MOVE_DO_MEM_READY: // check if all post init objects are finished with creating move DOs
      // if we're not in post init or the varan manager has finished waiting for post init objects => the move DO memory is ready
      if WaitForPostInitMoveObjectsCnt = 0 then
        pResult^.aData[4] := TRUE;
      else
        pResult^.aData[4] := FALSE;
      end_if;

//**********************************************************************************************************************************************************
    VM_CMD_SYNC_SEND_READY:
      // only work on it if the post init rt hasn't been finished, otherwise we would have the log messages if modules are plugged at runtime
      if b_PostInitRtSyncReady = FALSE then
        // Check Loader Version if function is supported
        if ops.uiLoaderVersion$UINT >= VM_POST_INIT_AVAILABLE then
          // only relevant during last Init
          if PostInitModuleCnt then
            // check if it's a valid index
            if pPara^.aPara[1]$UINT < VM_MAX_POST_INIT_MODULES then
              // check if our local this pointer matches this object
              if pPara^.aPara[0]$p_VaranBase = aPostInitList[pPara^.aPara[1]$UINT].p_This then
                // check if it's an object we were waiting for
                if aPostInitList[pPara^.aPara[1]$UINT].Settings.Wait4SyncSend then
                  aPostInitList[pPara^.aPara[1]$UINT].Settings.Wait4SyncSend := FALSE;

                  if WaitForSyncSendObjectsCnt then
                    WaitForSyncSendObjectsCnt -= 1;
                  else
#ifdef HWC_LogError
                    HWC_LogError(this, "@01B6 (VaranManager::Control::NewInst) There is already no more post init object to wait for (sync send ready)!");
#endif
                    ret_code := ERROR;
                  end_if;
                else
#ifdef HWC_LogError
                  HWC_LogError(this, "@01B7 (VaranManager::Control::NewInst) Module finished with sync send ready, where  There is already no more post init object to wait for!");
#endif
                  ret_code := ERROR;
                end_if;
              else
#ifdef HWC_LogError
                HWC_LogError(this, "@01B8 (VaranManager::Control::NewInst) This pointer of post init module given doesn't match locally stored this pointer for this index! (Move DOs)");
#endif
                ret_code := ERROR;
              end_if;
            else
#ifdef HWC_LogError
              HWC_LogError(this, "@01B9 (VaranManager::Control::NewInst) Invalid index of post init module given! (sync send ready)");
#endif
              ret_code := ERROR;
            end_if;
          else
#ifdef HWC_LogError
            HWC_LogError(this, "@01BA (VaranManager::Control::NewInst) More modules ready with last init than expected (sync send ready)");
#endif
            ret_code := ERROR;
          end_if;
        else
#ifdef HWC_LogError
          HWC_LogError(this, "@01B5 (VaranManager::Control::NewInst) VM_CMD_MOVE_DO_CREATION_FINISHED not supported with current Loader. Loader Version >= 02.02.137 is required (Move DOs)");
#endif
          ret_code := ERROR;
        end_if;
      end_if;

//**********************************************************************************************************************************************************
    VM_CMD_SET_MUX_THIS: // ignore this command, it's only for the VaranMux classes
      ret_code := ERROR; // return error => command not handled

//**********************************************************************************************************************************************************
    VM_CMD_INSTALL_DUMMY_CALLBACK:

      if pPara^.aPara[0] >= 4 * sizeof(DINT) then

        sd_retval := AddObjectCallback( p_us_position_info  := pPara^.aPara[1]$^USINT
                                      , ud_action_ptr       := pPara^.aPara[2]$UDINT
                                      , ud_thisp            := pPara^.aPara[3]$UDINT
                                      , sd_required         := pPara^.aPara[4]
                                      );
      else

#ifdef HWC_LogError
        HWC_LogError(this, "@01BB (VaranManager::Control::NewInst) VM_CMD_INSTALL_DUMMY_CALLBACK. Length of NewInst Commando is invalid");
#endif

      end_if;

//**********************************************************************************************************************************************************
    CMD_EXTEND_POST_INIT_TIME:
      // forward to HwControl
      To_HwControl.NewInst(pPara, pResult);

//**********************************************************************************************************************************************************
    CMD_GET_HW_TIMESTAMP:

      // forward to HwControl
      if pPara^.aPara[0]$t_GetHwTimestampCmd.udVersion = 1 then
        // Insert Coreselect if CmdVersion = 1 and increase CmdVersion to 2
        pPara^.aPara[0]$t_GetHwTimestampCmd.udVersion     := 2;
        pPara^.aPara[0]$t_GetHwTimestampCmd.udCoreSelect  := CoreSelect;
      end_if;
      ret_code := To_HwControl.NewInst(pPara, pResult);

//*****************************************************************************
    VM_CMD_GET_SYSTEM_MANAGER_CNT:

      pResult^.aData[0]$UDINT := udSystemVaranManagerCnt;

//**********************************************************************************************************************************************************
    CMD_HWC_REQ_PLLNS_REGULATION:
      // forward it to HwControl
      ret_code := To_HwControl.NewInst(pPara, pResult);

//**********************************************************************************************************************************************************
    else    // Commands for Payload
      if b_PayloadSupport then

        pResult^.uiLng          := sizeof(DINT);
        pResult^.aData[0]$DINT  := VM_CMD_NOT_IMPLEMENTED; // Default Return code, must be overwritten by induvidual methods

        CASE pPara^.uiCmd OF

        //*****************************************************************************
          VM_CMD_GET_MODULE_HANDLE :
            p_paraGetModuleHandel := (pPara^.aPara[0])$^t_VM_CMD_GetModuleHandle;

            pResult^.aData[0]$DINT := GetModuleHandle(  p_us_PositionInfo := p_paraGetModuleHandel^.p_us_position_info
                                                      , p_ud_ModuleHandle := p_paraGetModuleHandel^.p_ud_module_handle);

        //*****************************************************************************
          VM_CMD_ADD_DO :
            p_paraAddDO := (pPara^.aPara[0])$^t_VM_CMD_AddDO;
            pResult^.aData[0]$DINT := AddPayloadDO( p_ud_DoHandle                 := p_paraAddDO^.p_ud_DoHandle
                                                  , ud_NodeHandle                 := p_paraAddDO^.ud_ModuleHandle
                                                  , ud_DoRequired                 := p_paraAddDO^.ud_b_DoRequired
                                                  , ud_DolType                    := p_paraAddDO^.ud_DolType
                                                  , ud_Command                    := p_paraAddDO^.ud_Command
                                                  , ud_Priority                   := p_paraAddDO^.ud_Priority
                                                  , ud_PrescalerCounterThreshold  := p_paraAddDO^.ud_PreScalerCounterThreshold
                                                  , ud_PrescalerCounterStartValue := p_paraAddDO^.ud_PreScalerCounterStartValue
                                                  , ud_ReadOffset                 := p_paraAddDO^.ud_OffsetRead
                                                  , ud_ReadLength                 := p_paraAddDO^.ud_LengthRead
                                                  , ud_WriteOffset                := p_paraAddDO^.ud_OffsetWrite
                                                  , ud_WriteLength                := p_paraAddDO^.ud_LengthWrite
                                                  , ud_Filter                     := p_paraAddDO^.ud_Filter
                                                  , ud_Slices                     := p_paraAddDO^.ud_Slices
                                                  , ud_WritePayloadType           := p_paraAddDO^.ud_WritePayloadType);

        //*****************************************************************************
          VM_CMD_ADD_MOV_DO :
            p_paraMovDO := (pPara^.aPara[0])$^t_VM_CMD_AddMovDo;
            pResult^.aData[0]$DINT := AddPayloadMoveDO( p_ud_DoHandle                 := p_paraMovDO^.p_ud_DoHandle
                                                      , ud_bDoRequired                := p_paraMovDO^.ud_b_DoRequired
                                                      , ud_DolType                    := p_paraMovDO^.ud_DolType
                                                      , ud_Priority                   := p_paraMovDO^.ud_Priority
                                                      , ud_PrescalerCounterThreshold  := p_paraMovDO^.ud_PreScalerCounterThreshold
                                                      , ud_PrescalerCounterStartValue := p_paraMovDO^.ud_PreScalerCounterStartValue
                                                      , ud_hSourceReadDoHandle        := p_paraMovDO^.ud_SourceReadDoHandle
                                                      , ud_ReadOffset                 := p_paraMovDO^.ud_SourceReadOffset
                                                      , ud_hDestinationWriteDoHandle  := p_paraMovDO^.ud_DestinationWriteDoHandle
                                                      , ud_WriteOffset                := p_paraMovDO^.ud_DestinationWriteOffset
                                                      , ud_MoveDataLength             := p_paraMovDO^.ud_LengthMove);

        //*****************************************************************************
          VM_CMD_GET_DATA_POINTERS  :
            p_paraGetPointers := (pPara^.aPara[0])$^t_VM_CMD_GetDataPointers;
            pResult^.aData[0]$DINT := GetDataPointers(  ud_hDoHandle  := p_paraGetPointers^.ud_DoHandle
                                                      , pp_ReadData   := p_paraGetPointers^.p_ud_ReadData$^pVoid
                                                      , pp_WriteData  := p_paraGetPointers^.p_ud_WriteData$^pVoid);

        //*****************************************************************************
          VM_CMD_IS_DMA_ACTIVE :
            if PayloadFrame = 1 then
              pResult^.aData[0]$BOOL := TRUE;
            else
              pResult^.aData[0]$BOOL := FALSE;
            end_if;

        //*****************************************************************************
          else
            ret_code := ERROR;
        END_CASE;

      else
        pResult^.uiLng := sizeof(DINT);
        pResult^.aData[0]$DINT := VM_CMD_NOT_IMPLEMENTED;
#ifdef HWC_LogError
        HWC_LogError(this, "@01BC (VaranManager::Control::NewInst) Unknown command!");
#endif
        ret_code := ERROR;
      end_if;

  END_CASE;

END_FUNCTION

FUNCTION VaranManager::TurnOffIsoTask
  VAR
    s_PropertyValuePair : LSL_PROPERTY_VALUE_PAIR;
  END_VAR

  if b_PayloadSupport &
     pMultiVaran^.udVersion >= VM_MULTIVARAN_VERSION_FULL_PAYLOAD_AVAILABLE  then
    s_PropertyValuePair.udPropertyId    := VM_PROP_TASK_STATE_ISO;
    s_PropertyValuePair.udPropertyValue := TK_STATE_STOPPED;
    MULTI_VARAN_iSetNodeProperties( hNodeHandle           := vmNodeHandle
                                  , udPropertyCount       := 1
                                  , psPropertyValuePairs  := #s_PropertyValuePair
                                  );
  elsif p_ManagerStructure then
    p_ManagerStructure^.ucTCEnable := p_ManagerStructure^.ucTCEnable AND VM_DISABLE_ISO_TASK;
  end_if;

END_FUNCTION

FUNCTION VaranManager::AddPayloadDO
  VAR_INPUT
    p_ud_DoHandle 	                : ^UDINT;
    ud_NodeHandle 	                : UDINT;
    ud_DoRequired 	                : UDINT;
    ud_DolType 	                    : UDINT;
    ud_Command 	                    : UDINT;
    ud_Priority 	                  : UDINT;
    ud_PrescalerCounterThreshold 	  : UDINT;
    ud_PrescalerCounterStartValue 	: UDINT;
    ud_ReadOffset 	                : UDINT;
    ud_ReadLength 	                : UDINT;
    ud_WriteOffset 	                : UDINT;
    ud_WriteLength 	                : UDINT;
    ud_Filter 	  	                : UDINT;
    ud_Slices 	  	                : UDINT;
    ud_WritePayloadType             : UDINT;
  END_VAR
  VAR_OUTPUT
    sd_retval 	  	                : DINT;
  END_VAR
  VAR
    TempMem                         : UDINT;
    TempMemWr                       : UDINT;
  END_VAR

#ifdef VM_DEBUG_PAYLOAD
  if b_PayloadSupport = false then
    // This method is not suppored without payload
    ((0)$^USINT)^ := 0;
  end_if;
#endif

  //look if we Manager is on
  if ( ManagerOn ) then
    //look if we must execute Cyclic DOL list
    if ( ud_DolType = VARAN_DOL_ASY ) then
      s_CyHandles.b_ExecuteDOL := TRUE;			//set flag to execut Dol list
    end_if;

    sd_retval := MULTI_VARAN_iAddDo(  phDoHandle                    := p_ud_DoHandle
                                    , hNodeHandle                   := ud_NodeHandle
                                    , bDoRequired                   := ud_DoRequired
                                    , udDolType                     := ud_DolType
                                    , udCommand                     := ud_Command
                                    , udPriority                    := ud_Priority
                                    , udPrescalerCounterThreshold   := ud_PrescalerCounterThreshold
                                    , udPrescalerCounterStartValue  := ud_PrescalerCounterStartValue
                                    , udReadOffset                  := ud_ReadOffset
                                    , udReadLength                  := ud_ReadLength
                                    , udWriteOffset                 := ud_WriteOffset
                                    , udWriteLength                 := ud_WriteLength
                                    , udFilter                      := ud_Filter
                                    , udSlices                      := ud_Slices
                                    , udWritePayloadType            := ud_WritePayloadType$LSL_WRITE_PAYLOAD_TYPE);

    //look if an error occured
    if ( sd_retval <> VARANMANAGER_OK ) then
      s_ErrorVaranManager.f_AddRdDO := SetVaranDOError( sd_Error 		  := sd_retval
                                                      , b_manager_off	:= TRUE
                                                      , b_log			    := TRUE
                                                      );
    else

      if PayloadFrame = 1 then  // Use PayloadFrame because, b_PayloadSupport only shows the interface used.
                            // Payload DO Mem Calculaition +++++++++++++++++++++++++++++++++++++++++++++++++++++++++++++++++++++++++++++++++++++++++++++++++++++++++++++++++++++++++++++++++++++++++
        case ud_Command of

            VARAN_CMD_CONTROL_READ,
            VARAN_CMD_MEMORY_READ:      // Read DO -------------------------------------------------------------------------------------------------------------------------------
                // 1 Byte Status + n Byte (Load data read) + 0 to 3 Byte (compensate missalignment)
                TempMem := 1 + ud_ReadLength;

                // 1 Byte Control
                TempMemWr := 1;

                // Increase for variable DO
                if ud_WritePayloadType > WR_PLD_TYPE_STANDARD$UDINT then
                  TempMemWr += 16#0E;
                end_if;

                case ud_DolType of
                // **************************************************
                  VARAN_DOL_DA:
                    DPRAM_Used.DA_Rd            += TempMem + TempMemWr + SIZE_PAYLOAD_FRAME_HEADER_DO;
                    DPRAM_Used_Payload.DA_Rd    += TempMem;
                    DPRAM_Used_Payload.DA_Wr    += TempMemWr;
                    DOCounter.DA_Rd             += 1;

                // **************************************************
                  VARAN_DOL_ISO:
                    DPRAM_Used.ISO_Rd           += TempMem + TempMemWr + SIZE_PAYLOAD_FRAME_HEADER_DO;
                    DPRAM_Used_Payload.ISO_Rd   += TempMem;
                    DPRAM_Used_Payload.ISO_Wr   += TempMemWr;
                    DOCounter.ISO_Rd            += 1;

                // **************************************************
                  VARAN_DOL_ASY:
                    DPRAM_Used.ASY_Rd           += TempMem + TempMemWr + SIZE_PAYLOAD_FRAME_HEADER_DO;
                    DPRAM_Used_Payload.ASY_Rd   += TempMem;
                    DPRAM_Used_Payload.ASY_Wr   += TempMemWr;
                    DOCounter.ASY_Rd            += 1;

                // **************************************************
                  VARAN_DOL_ADMIN:
                    DPRAM_Used.Admin_Rd         += TempMem + TempMemWr + SIZE_PAYLOAD_FRAME_HEADER_DO;
                    DPRAM_Used_Payload.Admin_Rd += TempMem;
                    DPRAM_Used_Payload.ASY_Wr   += TempMemWr;
                    DOCounter.Admin_Rd          += 1;

                // **************************************************
                  VARAN_DOL_IRQ:
                    DPRAM_Used.IRQ_Rd         += TempMem + TempMemWr + SIZE_PAYLOAD_IRQ_FRAME_HEADER_DO;
                    DPRAM_Used_Payload.IRQ_Rd += TempMem;
                    DPRAM_Used_Payload.IRQ_Wr += TempMemWr;
                    DOCounter.IRQ_Rd          += 1;
                end_case;

                DPRAM_Used_Payload.Payload_Read     += TempMem;
                DPRAM_Used_Payload.Payload_Write    += TempMemWr;

                if ud_DolType <> VARAN_DOL_IRQ then
                  DPRAM_Used.Total                  += TempMem + TempMemWr + SIZE_PAYLOAD_FRAME_HEADER_DO;
                  DPRAM_Used_Payload.Payload_Header += SIZE_PAYLOAD_FRAME_HEADER_DO;
                else
                  DPRAM_Used.Total                  += TempMem + TempMemWr + SIZE_PAYLOAD_IRQ_FRAME_HEADER_DO;
                  DPRAM_Used_Payload.Payload_Header += SIZE_PAYLOAD_IRQ_FRAME_HEADER_DO;
                end_if;

                DPRAM_Used_Payload.Total            += TempMem + TempMemWr;

                DOCounter.Total                     += 1;

            VARAN_CMD_CONTROL_WRITE,
            VARAN_CMD_MEMORY_WRITE:     // Write DO -------------------------------------------------------------------------------------------------------------------------------
                // 1 Byte Control + n Byte (Load data read) + 0 to 3 Byte (compensate missalignment)
                TempMemWr := 1 + ud_WriteLength;

                // Increase for variable DO
                if ud_WritePayloadType > WR_PLD_TYPE_STANDARD$UDINT then
                  TempMemWr += 16#0E;
                end_if;

                // 1 Byte Status in Read DPRAM
                TempMem := 1;

                case ud_DolType of
                // **************************************************
                  VARAN_DOL_DA:
                    DPRAM_Used.DA_Wr            += TempMem + TempMemWr + SIZE_PAYLOAD_FRAME_HEADER_DO;
                    DPRAM_Used_Payload.DA_Rd    += TempMem;
                    DPRAM_Used_Payload.DA_Wr    += TempMemWr;
                    DOCounter.DA_Wr             += 1;

                // **************************************************
                  VARAN_DOL_ISO:
                    DPRAM_Used.ISO_Wr           += TempMem + TempMemWr + SIZE_PAYLOAD_FRAME_HEADER_DO;
                    DPRAM_Used_Payload.ISO_Rd   += TempMem;
                    DPRAM_Used_Payload.ISO_Wr   += TempMemWr;
                    DOCounter.ISO_Wr            += 1;

                // **************************************************
                  VARAN_DOL_ASY:
                    DPRAM_Used.ASY_Wr           += TempMem + TempMemWr + SIZE_PAYLOAD_FRAME_HEADER_DO;
                    DPRAM_Used_Payload.ASY_Rd   += TempMem;
                    DPRAM_Used_Payload.ASY_Wr   += TempMemWr;
                    DOCounter.ASY_Wr            += 1;

                // **************************************************
                  VARAN_DOL_ADMIN:
                    DPRAM_Used.Admin_Wr         += TempMem + TempMemWr + SIZE_PAYLOAD_FRAME_HEADER_DO;
                    DPRAM_Used_Payload.Admin_Rd += TempMem;
                    DPRAM_Used_Payload.Admin_Wr += TempMemWr;
                    DOCounter.Admin_Wr          += 1;

                // **************************************************
                  VARAN_DOL_IRQ:
                    DPRAM_Used.IRQ_Wr           += TempMem + TempMemWr + SIZE_PAYLOAD_IRQ_FRAME_HEADER_DO;
                    DPRAM_Used_Payload.ISO_Rd   += TempMem;
                    DPRAM_Used_Payload.IRQ_Wr   += TempMemWr;
                    DOCounter.IRQ_Wr            += 1;

                end_case;

                DPRAM_Used_Payload.Payload_Read     += TempMem;
                DPRAM_Used_Payload.Payload_Write    += TempMemWr;

                if ud_DolType <> VARAN_DOL_IRQ then
                  DPRAM_Used.Total                  += TempMem + TempMemWr + SIZE_PAYLOAD_FRAME_HEADER_DO;
                  DPRAM_Used_Payload.Payload_Header += SIZE_PAYLOAD_FRAME_HEADER_DO;
                else
                  DPRAM_Used.Total                  += TempMem + TempMemWr + SIZE_PAYLOAD_IRQ_FRAME_HEADER_DO;
                  DPRAM_Used_Payload.Payload_Header += SIZE_PAYLOAD_IRQ_FRAME_HEADER_DO;
                end_if;

                DPRAM_Used_Payload.Total            += TempMem + TempMemWr;
                DOCounter.Total                     += 1;

            VARAN_CMD_CONTROL_READ_WRITE,
            VARAN_CMD_MEMORY_READ_WRITE:// Read/Write DO -------------------------------------------------------------------------------------------------------------------------------
                // 1 Byte Control + n Byte (Load data read) + 0 to 3 Byte (compensate missalignment) x2
                TempMem   := 1 + ud_ReadLength;

                TempMemWr := 1 + ud_WriteLength;

                // Increase for variable DO
                if ud_WritePayloadType = WR_PLD_TYPE_RW_ACCESS_CONFIGURABLE$UDINT then
                  TempMemWr += 16#14;
                elsif ud_WritePayloadType > WR_PLD_TYPE_STANDARD$UDINT then
                  TempMemWr += 16#0E;
                end_if;

                case ud_DolType of
                // **************************************************
                  VARAN_DOL_DA:
                    DPRAM_Used.DA_RdWr          += TempMem + TempMemWr + SIZE_PAYLOAD_FRAME_HEADER_DO;
                    DPRAM_Used_Payload.DA_Rd    += TempMem;
                    DPRAM_Used_Payload.DA_Wr    += TempMemWr;
                    DOCounter.DA_RdWr           += 1;

                // **************************************************
                  VARAN_DOL_ISO:
                    DPRAM_Used.ISO_RdWr         += TempMem + TempMemWr + SIZE_PAYLOAD_FRAME_HEADER_DO;
                    DPRAM_Used_Payload.ISO_Rd   += TempMem;
                    DPRAM_Used_Payload.ISO_Wr   += TempMemWr;
                    DOCounter.ISO_RdWr          += 1;

                // **************************************************
                  VARAN_DOL_ASY:
                    DPRAM_Used.ASY_RdWr         += TempMem + TempMemWr + SIZE_PAYLOAD_FRAME_HEADER_DO;
                    DPRAM_Used_Payload.ASY_Rd   += TempMem;
                    DPRAM_Used_Payload.ASY_Wr   += TempMemWr;
                    DOCounter.ASY_RdWr          += 1;

                // **************************************************
                  VARAN_DOL_ADMIN:
                    DPRAM_Used.Admin_RdWr       += TempMem + TempMemWr + SIZE_PAYLOAD_FRAME_HEADER_DO;
                    DPRAM_Used_Payload.Admin_Rd += TempMem;
                    DPRAM_Used_Payload.Admin_Wr += TempMemWr;
                    DOCounter.Admin_RdWr        += 1;

                // **************************************************
                  VARAN_DOL_IRQ:
                    DPRAM_Used.IRQ_RdWr         += TempMem + TempMemWr + SIZE_PAYLOAD_IRQ_FRAME_HEADER_DO;
                    DPRAM_Used_Payload.IRQ_Rd   += TempMem;
                    DPRAM_Used_Payload.IRQ_Wr   += TempMemWr;
                    DOCounter.IRQ_RdWr          += 1;

                end_case;

                DPRAM_Used_Payload.Payload_Read     += TempMem;
                DPRAM_Used_Payload.Payload_Write    += TempMemWr;

                if ud_DolType <> VARAN_DOL_IRQ then
                  DPRAM_Used.Total                  += TempMem + TempMemWr + SIZE_PAYLOAD_FRAME_HEADER_DO;
                  DPRAM_Used_Payload.Payload_Header += SIZE_PAYLOAD_FRAME_HEADER_DO;
                else
                  DPRAM_Used.Total                  += TempMem + TempMemWr + SIZE_PAYLOAD_IRQ_FRAME_HEADER_DO;
                  DPRAM_Used_Payload.Payload_Header += SIZE_PAYLOAD_IRQ_FRAME_HEADER_DO;
                end_if;

                DPRAM_Used_Payload.Total            += TempMem + TempMemWr;
                DOCounter.Total                     += 1;

        end_case;
      else    // Standard DO Mem Calculation +++++++++++++++++++++++++++++++++++++++++++++++++++++++++++++++++++++++++++++++++++++++++++++++++++++++++++++++++++++++++++++++++++++++++

        case ud_Command of

            VARAN_CMD_CONTROL_READ,
            VARAN_CMD_MEMORY_READ:      // Read DO -------------------------------------------------------------------------------------------------------------------------------
                // 32 Byte (Header) + 6 Byte (1 Byte Cmd, 4 Byte Addr, 1 Byte Len) + 1 Byte (Response) + n Byte (Load data read) + 0 to 3 Byte (compensate missalignment)
                TempMem := 32 + 6 + 1 + ud_ReadLength;
                if (TempMem MOD 4) then
                  TempMem := TempMem + (4 - (TempMem MOD 4)); //increase memory, up to a value, which could be divided by 4
                end_if;

                case ud_DolType of
                // **************************************************
                  VARAN_DOL_DA:
                                DPRAM_Used.DA_Rd    += TempMem;
                                DOCounter.DA_Rd     += 1;
                // **************************************************
                  VARAN_DOL_ISO:
                                DPRAM_Used.ISO_Rd   += TempMem;
                                DOCounter.ISO_Rd    += 1;
                // **************************************************
                  VARAN_DOL_ASY:
                                DPRAM_Used.ASY_Rd   += TempMem;
                                DOCounter.ASY_Rd    += 1;
                // **************************************************
                  VARAN_DOL_ADMIN:
                                DPRAM_Used.Admin_Rd += TempMem;
                                DOCounter.Admin_Rd  += 1;
                // **************************************************
                  VARAN_DOL_IRQ:
                                DPRAM_Used.IRQ_Rd   += TempMem;
                                DOCounter.IRQ_Rd    += 1;
                end_case;

                DPRAM_Used.Total  += TempMem;
                DOCounter.Total   += 1;

            VARAN_CMD_CONTROL_WRITE,
            VARAN_CMD_MEMORY_WRITE:     // Write DO -------------------------------------------------------------------------------------------------------------------------------
                //32 Byte (Header) + 6 Byte (1 Byte Cmd, 4 Byte Addr, 1 Byte Len) + 1 Byte (Response) + n Byte (load data write) + 0 to 3 Byte (compensate missalignment)
                  TempMem := 32 + 6 + 1 + ud_WriteLength;
                  if (TempMem MOD 4) then
                    TempMem := TempMem + (4 - (TempMem MOD 4)); //increase memory, up to a value, which could be divided by 4
                  end_if;

                  case ud_DolType of
                  // **************************************************
                    VARAN_DOL_DA:
                                  DPRAM_Used.DA_Wr    += TempMem;
                                  DOCounter.DA_Wr     += 1;
                  // **************************************************
                    VARAN_DOL_ISO:
                                  DPRAM_Used.ISO_Wr   += TempMem;
                                  DOCounter.ISO_Wr    += 1;
                  // **************************************************
                    VARAN_DOL_ASY:
                                  DPRAM_Used.ASY_Wr   += TempMem;
                                  DOCounter.ASY_Wr    += 1;
                  // **************************************************
                    VARAN_DOL_ADMIN:
                                  DPRAM_Used.Admin_Wr += TempMem;
                                  DOCounter.Admin_Wr  += 1;
                  // **************************************************
                    VARAN_DOL_IRQ:
                                  DPRAM_Used.IRQ_Wr   += TempMem;
                                  DOCounter.IRQ_Wr    += 1;
                  end_case;

                  DPRAM_Used.Total  += TempMem;
                  DOCounter.Total   += 1;

            VARAN_CMD_CONTROL_READ_WRITE,
            VARAN_CMD_MEMORY_READ_WRITE:// Read/Write DO -------------------------------------------------------------------------------------------------------------------------------
                  //32 Byte (Header) + 11 Byte (1 Byte Cmd, 4 Byte RdAddr, 1 Byte RdLen, 4 Byte WrAddr, 1 Byte WrLen) + 1 Byte (Response) + n Byte (load data read) + n Byte (load data write) + 0 to 3 Byte (compensate missalignment)
                  TempMem := 32 + 11 + 1 + ud_ReadLength + ud_WriteLength;
                  if (TempMem MOD 4) then
                    TempMem := TempMem + (4 - (TempMem MOD 4)); //increase memory, up to a value, which could be divided by 4
                  end_if;

                  case ud_DolType of
                  // **************************************************
                    VARAN_DOL_DA:
                                  DPRAM_Used.DA_RdWr    += TempMem;
                                  DOCounter.DA_RdWr     += 1;
                  // **************************************************
                    VARAN_DOL_ISO:
                                  DPRAM_Used.ISO_RdWr   += TempMem;
                                  DOCounter.ISO_RdWr    += 1;
                  // **************************************************
                    VARAN_DOL_ASY:
                                  DPRAM_Used.ASY_RdWr   += TempMem;
                                  DOCounter.ASY_RdWr    += 1;
                  // **************************************************
                    VARAN_DOL_ADMIN:
                                  DPRAM_Used.Admin_RdWr += TempMem;
                                  DOCounter.Admin_RdWr  += 1;
                  // **************************************************
                    VARAN_DOL_IRQ:
                                  DPRAM_Used.IRQ_RdWr   += TempMem;
                                  DOCounter.IRQ_RdWr    += 1;
                  end_case;

                  DPRAM_Used.Total  += TempMem;
                  DOCounter.Total   += 1;

        end_case;

      end_if; // +++++++++++++++++++++++++++++++++++++++++++++++++++++++++++++++++++++++++++++++++++++++++++++++++++++++++++++++++++++++++++++++++++++++++++++++++++++++++++++++++++++++++++++++++

    end_if;
  else
    sd_retval := -100;	//Manager is off
  end_if;
END_FUNCTION

FUNCTION VaranManager::AddPayloadMoveDO
  VAR_INPUT
    p_ud_DoHandle 	                : ^UDINT;
    ud_bDoRequired 	                : UDINT;
    ud_DolType 	                    : UDINT;
    ud_Priority 	                  : UDINT;
    ud_PrescalerCounterThreshold 	  : UDINT;
    ud_PrescalerCounterStartValue 	: UDINT;
    ud_hSourceReadDoHandle 	        : UDINT;
    ud_ReadOffset 	                : UDINT;
    ud_hDestinationWriteDoHandle 	  : UDINT;
    ud_WriteOffset 	                : UDINT;
    ud_MoveDataLength 	            : UDINT;
  END_VAR
  VAR_OUTPUT
    sd_retval 	                    : DINT;
  END_VAR

#ifdef VM_DEBUG_PAYLOAD
  if b_PayloadSupport = false then
    // This method is not suppored without payload
    ((0)$^USINT)^ := 0;
  end_if;
#endif

  //look if we must execute Cyclic DOL list
  if ( ud_DolType = VARAN_DOL_ASY ) then
    s_CyHandles.b_ExecuteDOL := TRUE;			//set flag to execut Dol list
  end_if;

  sd_retval := MULTI_VARAN_iAddMoveDo(  phDoHandle                    := p_ud_DoHandle
                                      , bDoRequired                   := ud_bDoRequired
                                      , udDolType                     := ud_DolType
                                      , udPriority                    := ud_Priority
                                      , udPrescalerCounterThreshold   := ud_PrescalerCounterThreshold
                                      , udPrescalerCounterStartValue  := ud_PrescalerCounterStartValue
                                      , hSourceReadDoHandle           := ud_hSourceReadDoHandle
                                      , udReadOffset                  := ud_ReadOffset
                                      , hDestinationWriteDoHandle     := ud_hDestinationWriteDoHandle
                                      , udWriteOffset                 := ud_WriteOffset
                                      , udMoveDataLength              := ud_MoveDataLength
                                      );
  //look if an error occured
  if ( sd_retval <> VARANMANAGER_OK ) then
    s_ErrorVaranManager.f_AddRdDO := SetVaranDOError( sd_Error      := sd_retval
                                                    , b_manager_off := TRUE
                                                    , b_log         := TRUE
                                                    );
  else
    // Payload Move DO Mem Calculation
    if ( ud_DolType = VARAN_DOL_ASY ) then
      DPRAM_Used.ASY_Mov          += sizeof(LSL_VARANFRAMEPAYLOADMOVEHEADER);
      DPRAM_Used_Payload.ASY_Rd   += 1; // 1 Byte status
      DPRAM_Used_Payload.ASY_Wr   += sizeof(LSL_VARANFRAMEMOVEWRITEPAYLOAD);
      DOCounter.ASY_Mov           += 1;
    else
      DPRAM_Used.ISO_Mov          += sizeof(LSL_VARANFRAMEPAYLOADMOVEHEADER);
      DPRAM_Used_Payload.ISO_Rd   += 1; // 1 Byte status
      DPRAM_Used_Payload.ISO_Wr   += sizeof(LSL_VARANFRAMEMOVEWRITEPAYLOAD);
      DOCounter.ISO_Mov           += 1;
    end_if;
